PROGRAM Control_FBD
VAR
	ixSensor1		AT %I*:	BOOL; 		//Pallet on sensor1 (S1)
	ixSensor2		AT %I*:	BOOL; 		//Pallet on sensor2 (S2)
	ixSensor3		AT %I*:	BOOL; 		//Pallet on sensor3 (S3)

	qxRunConveyor1	AT %Q*:	BOOL; 		// Motor that runs Conveyor 1*)
	qxRunConveyor2	AT %Q*:	BOOL; 		// Motor that runs Conveyor 2*)
	qxRunConveyor3	AT %Q*:	BOOL; 		// Motor that runs Conveyor 3*)	

	//Transport memory
	mxTrpConveyor1to2 : BOOL;
	mxTrpConveyor2to3 : BOOL;

END_VAR

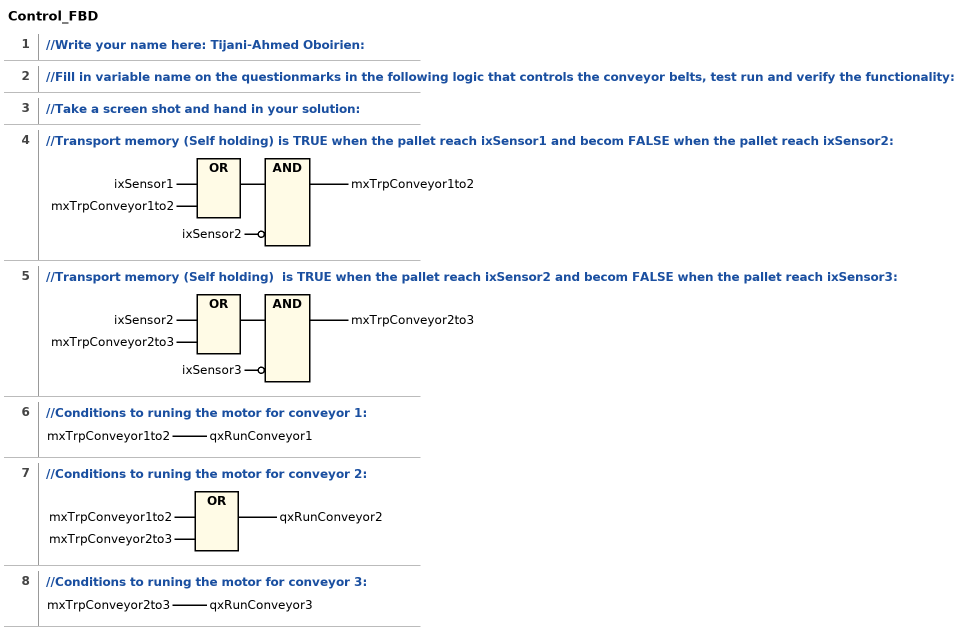
// NETWORK 1
// label: //Write your name here: Tijani-Ahmed Oboirien

// NETWORK 2
// label: //Fill in variable name on the questionmarks in the following logic that controls the conveyor belts, test run and verify the functionality

// NETWORK 3
// label: //Take a screen shot and hand in your solution

// NETWORK 4
// label: //Transport memory (Self holding) is TRUE when the pallet reach ixSensor1 and becom FALSE when the pallet reach ixSensor2
mxTrpConveyor1to2 := (ixSensor1 OR mxTrpConveyor1to2) AND NOT ixSensor2;

// NETWORK 5
// label: //Transport memory (Self holding)  is TRUE when the pallet reach ixSensor2 and becom FALSE when the pallet reach ixSensor3
mxTrpConveyor2to3 := (ixSensor2 OR mxTrpConveyor2to3) AND NOT ixSensor3;

// NETWORK 6
// label: //Conditions to runing the motor for conveyor 1
qxRunConveyor1 := mxTrpConveyor1to2;

// NETWORK 7
// label: //Conditions to runing the motor for conveyor 2
qxRunConveyor2 := mxTrpConveyor1to2 OR mxTrpConveyor2to3;

// NETWORK 8
// label: //Conditions to runing the motor for conveyor 3
qxRunConveyor3 := mxTrpConveyor2to3;

END_PROGRAM

(* stored: Version 1.1.0.1
   POU Control_FBD: Id {84d3f40d-a0f6-423e-bc58-eeabb716185d}, SpecialFunc None *)
